Fanuc KAREL source: kt00153.KL

-- PROVISIONAL review KL for V770-1; original PC SHA256 7538a6b7d6c12aae4b9875fe339d11045f13f66c7e680f9efbc2de34e6e02d55
-- Incomplete behavior may be omitted. Consult companion uncertainty JSON. Do not deploy.
PROGRAM KT00153
%NOLOCKGROUP
VAR
  I2 : INTEGER
  OUT : INTEGER
-- UNRESOLVED_DECL H1 type=002017
BEGIN
  -- UNRESOLVED_PC offsets 5-19; opcodes 2E,22,9D,33,B4
  -- UNRESOLVED_PC offsets 24-35; opcodes 2E,23
  -- UNRESOLVED_PC offsets 40-62; opcodes 22,9D,33,B3,21,55,23
  -- UNRESOLVED_PC offsets 67-71; opcodes 7F
END KT00153
